(* IEC 61131-3 sources: JingjiangArm/moonboxpro_arm_8.4/Application/Application/任务列表/Main_Task/套色调整/套色新算法/PID_GET, 9 files *)

(* ---- AntiNotch_1.st ---- *)
(*@CES
Name=AntiNotch_1
Type=FunctionBlock
TypeGuid=6f9dac99-8de1-4efc-8465-68ac443b7d08
Guid=fc76d1c1-3b33-4f49-ab68-3746014dafce
HasDeclaration=True
HasImplementation=True
*)
{DECLARATION}
FUNCTION AntiNotch_1 : BOOL
(*功能：反陷波器(s^2+2*d*wn*s+wn^2)/(s^2+2*d*xi*wn*s+wn^2)的差分方程实现*)
(*输入：*)
(*输出：*)
VAR_INPUT
	i_rU:REAL;(*信号输入*)
	i_prYout: POINTER TO REAL;(*信号输出*)

(*(s^2+2*d*wn*s+wn^2)/(s^2+2*d*xi*wn*s+wn^2)*)
	i_rWn:REAL;(*陷波中心频率 rad/s*)
	i_rBw:REAL;(*陷波宽度 rad/s*)
	i_rDp:REAL;(*陷波深度 dB*)

	i_rTs:REAL;(*采样时间*)

	i_prUk:POINTER TO ARRAY [1..3] OF REAL;(*输入寄存器*)
	i_prYk:POINTER TO ARRAY [1..3] OF REAL;(*输出寄存器*)
END_VAR
VAR
	rFn:REAL:=0;
	rFBw:REAL:=0;
	rWn:REAL:=0;
	rDp:REAL:=0;

	rD:REAL:=0;
	rXi:REAL:=0;

	rK:REAL:=0;
	ra2:REAL:=0;
	ra1:REAL:=0;
	ra0:REAL:=0;

	rb2:REAL:=0;
	rb1:REAL:=0;
	rb0:REAL:=0;

	rTs:REAL:=0;(*采样时间*)
	rTemp:REAL:=0;

END_VAR
{IMPLEMENTATION}
(*参数初始化*)
rFn := i_rWn/2.0*gc_lrPi;
rWn := i_rWn;
rFBw := i_rBw/2.0*gc_lrPi;
rDp := i_rDp;

rTemp := -rDp/20.0;
rD := EXPT(10,rTemp);

rTemp := 1.0/(1.0 - 2.0*EXPT(rD,2));
rXi := rFBw/(2.0*rFn)*SQRT(rTemp);

rK := 1.0;

ra2:=1.0;
ra1:=2*rXi*rWn;
ra0:=rWn*rWn;

rb2:=1;
rb1:=2*rD*rXi*rWn;
rb0:=rWn*rWn;

rTs:=i_rTs;

(*更新寄存器注意顺序*)
i_prYk^[3]:=i_prYk^[2];
i_prYk^[2]:=i_prYk^[1];

i_prUk^[3]:=i_prUk^[2];
i_prUk^[2]:=i_prUk^[1];

(*差分计算*)
i_prUk^[1]:=rK*i_rU;
rTemp:=1/(rb0*rTs*rTs+2*rb1*rTs+4*rb2)*(-(2*rb0*rTs*rTs-8*rb2)*i_prYk^[2]-(rb0*rTs*rTs-2*rb1*rTs+4*rb2)*i_prYk^[3]
            +(ra0*rTs*rTs+2*ra1*rTs+4*ra2)*i_prUk^[1]+(2*ra0*rTs*rTs-8*ra2)*i_prUk^[2]+(ra0*rTs*rTs-2*ra1*rTs+4*ra2)*i_prUk^[3]);
i_prYk^[1]:=rTemp;
i_prYout^:=rTemp;

(* ---- Cal_Kp_Ki.st ---- *)
(*@CES
Name=Cal_Kp_Ki
Type=FunctionBlock
TypeGuid=6f9dac99-8de1-4efc-8465-68ac443b7d08
Guid=a93d564e-2599-4b4b-9c00-c963b5a75637
HasDeclaration=True
HasImplementation=True
*)
{DECLARATION}
FUNCTION Cal_Kp_Ki : BOOL
(*2024.9.6.123503*)
(*通过和控制器计算公式对比这里对Ki做的一些处理,反应到Ki计算上相当于积分的系数是定值,因为ts=周长/速度*系数
这里对输入的i_rV 按照30m/min定值输入,这样在计算积分的时候会出现积分根据速度逐渐减小的变化*)
(*2024.9.6.125139 将Ki的速度分开*)
(*2025.1.3.140421删除无用的*)
VAR_INPUT
(*
	i_byFilmType:BYTE;
	(*增加一些控制变量@2024.8.25.164242*)
	i_byTimingKiByArcErr:BYTE;(*=0 不使能|=1根据误差值Ki变化|值越大积分越小*)
	i_byAverageNum:BYTE;(*平均次数*)
	i_byColorId:BYTE;(*色序id*)
	i_iArcErr:INT;(*套色误差@mm*)
*)
(*模型变量*)
	i_rV:REAL;(*运行速度m/min*)
	i_rV_Ki:REAL;(*运行速度m/min*)
	i_rCL:REAL;(*版周长mm*)
	i_rL:REAL;(*机组料长m*)
(*控制变量*)
	i_rKadj_all:REAL;(*调整增益   40*)
	i_rKadj_i:REAL;(*积分增益  2.0*)
(*输出指针*)
	i_prKp:POINTER TO REAL;(*Kp*)
	i_prKi:POINTER TO REAL;(*Ki*)
END_VAR
VAR

	rA:REAL;(*模型参数*)(*
	iAverageNum:INT;
	iArcErr:INT;
*)
END_VAR
{IMPLEMENTATION}
IF i_rL<>0 AND i_rV<>0 AND i_rV_Ki<>0 AND i_rCL<>0 THEN
	(*计算模型参数*)
	rA := (i_rV/60.0)/i_rL;
	(*Kp*)
	i_prKp^ := i_rKadj_all/i_rCL*i_rV/rA;

	(*Ki*)
(*	i_prKi^ := i_rKadj_all/i_rCL*i_rV*i_rKadj_i;*)
	i_prKi^ := i_rKadj_all/i_rCL*i_rV_Ki*i_rKadj_i;
ELSE
	i_prKp^ := 16;
	i_prKi^ := 8;
END_IF

(* ---- Cal_Kp_Ki_V2.st ---- *)
(*@CES
Name=Cal_Kp_Ki_V2
Type=FunctionBlock
TypeGuid=6f9dac99-8de1-4efc-8465-68ac443b7d08
Guid=c47de549-0752-4bbe-8145-8113c580532b
HasDeclaration=True
HasImplementation=True
*)
{DECLARATION}
FUNCTION Cal_Kp_Ki_V2 : BOOL
(*2025.1.15.123422 增加了时延参数输入*)
VAR_INPUT
(*模型变量*)
	i_rV:REAL;(*运行速度m/min*)
	i_rLTao:REAL;(*印刷点到光电眼距离*)
	i_rL:REAL;(*机组料长m*)
	i_rDelay:REAL;(*时延@2025.1.15.123404+*)
(*控制变量*)
	i_rKadj_Mag:REAL;(*幅值裕度   15dB|越小越强*)
	i_rKadj_i:REAL;(*积分增益  1.0*)
(*输出指针*)
	i_prKp:POINTER TO REAL;(*Kp*)
	i_prKi:POINTER TO REAL;(*Ki*)
END_VAR
VAR
	rA:REAL;(*模型参数*)
	rTao:REAL;(*光电眼到印刷点的时延 s*)

	rWf:REAL;(*-180度对应的频率*)
	rMag_Wf:REAL;(*-180度对应的幅值*)

	rKadj:REAL; (*满足幅值裕度的增益*)
	rKTemp:REAL;(*增益计算临时变量*)

	iAverageNum:INT;
	iArcErr:INT;
END_VAR
{IMPLEMENTATION}
IF i_rL<>0 AND i_rV<>0 AND i_rLTao<>0 THEN
	(*计算模型参数*)
	rA := (i_rV/60.0)/i_rL;
(*	rTao := i_rLTao/(i_rV/60.0) +0.1 ;*)
	rTao := i_rLTao/(i_rV/60.0) + i_rDelay ;

	(*计算-180度对应的频率*)
	rWf := LREAL_TO_REAL(90.0 * gc_lrPi / 180.0 / rTao);
	(*计算-180度对应的幅值 和rKadj*)
	rMag_Wf := 20.0 * LOG(0.1 * rA / rWf); (*为负数*)
	rKTemp := (-1.0*i_rKadj_Mag - rMag_Wf) / 20.0  ;
	rKadj := LREAL_TO_REAL(EXPT(10, rKTemp));

	(*Kp*)
	i_prKp^ := rKadj;

	(*Ki*)
	i_prKi^ := rKadj * rA * i_rKadj_i;
ELSE
	i_prKp^ := 16;
	i_prKi^ := 8;
END_IF

(* ---- Cal_Kp_Ki_V3.st ---- *)
(*@CES
Name=Cal_Kp_Ki_V3
Type=FunctionBlock
TypeGuid=6f9dac99-8de1-4efc-8465-68ac443b7d08
Guid=deaeaf1e-1ab7-4a2c-8f0b-a36d361ddac8
HasDeclaration=True
HasImplementation=True
*)
{DECLARATION}
FUNCTION Cal_Kp_Ki_V3 : BOOL
(*2025.1.11.165519 增加了非法值处理@Liu.yt*)
(*将开环对象镇定为期望的幅值裕度和相位裕度*)
(*输入开环幅值裕度(10-20)，相位裕度(40-60)*)
(*由于需要调整积分满足相位裕度，因此实际的幅值裕度会略微小于设置值（在所给出的相位裕度范围内一般偏差在1dB以内，不超过2dB），相位裕度取得越小，幅值裕度偏差越大*)

VAR_INPUT
(*模型变量*)
	i_rV:REAL;(*运行速度m/min*)
	i_rLTao:REAL;(*印刷点到光电眼距离*)
	i_rL:REAL;(*机组料长m*)
(*控制变量*)
	i_rMargin_Mag:REAL;(*幅值裕度   15dB*)
	i_rMargin_Phi:REAL;(*相位裕度  50度*)
(*输出指针*)
	i_prKp:POINTER TO REAL;(*Kp*)
	i_prKi:POINTER TO REAL;(*Ki*)
END_VAR
VAR
	rA:REAL;(*模型参数*)
	rTao:REAL;(*光电眼到印刷点的时延 s*)

	rWf:REAL;(*-180度对应的频率*)
	rMag_Wf:REAL;(*-180度对应的幅值*)

	rKadj:REAL; (*满足幅值裕度的增益*)
	rKTemp:REAL;(*增益计算临时变量*)

	rKp_temp:REAL; (*临时Kp*)
	rKi_temp:REAL;(*临时Ki*)

	rax:REAL; (*模型临时参数，计算Wc使用*)
	rbx:REAL; (*模型临时参数，计算Wc使用*)

	rA_e:REAL;(*二次方程系数*)
	rB_e:REAL;(*二次方程系数*)
	rC_e:REAL;(*二次方程系数*)

	rX_temp:REAL;(*方程的解*)
	rWc:REAL;(*近似截止频率*)

	rPhi_temp:REAL;(*相位裕度临时量*)
	rDelta_Phi:REAL;(*相位裕度偏差*)
	rDelta_Phi_rad:REAL;(*相位裕度偏差 弧度表示*)

	rI:REAL;(*积分系数*)
END_VAR
{IMPLEMENTATION}
IF i_rL<>0 AND i_rV<>0 AND i_rLTao<>0 THEN
(*计算模型参数*)
	rA := (i_rV/60.0)/i_rL;
	rTao := i_rLTao/(i_rV/60.0) +0.1 ;
(*计算满足幅值裕度时的近似截止频率和增益*)
	(*计算-180度对应的频率*)
	rWf := LREAL_TO_REAL(90.0 * gc_lrPi / 180.0 / rTao);
	(*计算-180度对应的幅值 和rKadj*)
	rMag_Wf := 20.0 * LOG(0.1 * rA / rWf); (*为负数*)
	rKTemp := (-1.0*i_rMargin_Mag - rMag_Wf) / 20.0  ;
	rKadj := LREAL_TO_REAL(EXPT(10, rKTemp));

	(*Kp*)
	rKp_temp := rKadj;

	(*Ki*)
	rKi_temp := rKadj * rA;
	(*计算此时的截止频率Wc*)
	rax := rA;
	rbx := 0.1*rA;

	(*构建二次方程*)
	rA_e := 1;
	rB_e := rax * rax - rbx * rbx * rKp_temp * rKp_temp;
	rC_e := -1.0 * rbx * rbx * rKi_temp * rKi_temp;

	(*计算根*)
	rX_temp := (-1.0 * rB_e + SQRT(rB_e * rB_e - 4.0 * rA_e * rC_e)) / (2.0 * rA_e);
	rWc := SQRT(rX_temp);

	(*计算相位裕度偏差*)
	rPhi_temp := LREAL_TO_REAL(90.0 - rWc * rTao / gc_lrPi * 180.0);
	rDelta_Phi := rPhi_temp - i_rMargin_Phi - 5;(*5是额外的裕度，可调整*)

	rI := rA;
	IF rDelta_Phi > 0 THEN
		(*转成弧度表示*)
		rDelta_Phi_rad := LREAL_TO_REAL(rDelta_Phi / 180.0 * gc_lrPi);

		(*计算调整的积分系数rI *)
		rI := rWc * (1.0 + (rWc / rA) * TAN(rDelta_Phi_rad) ) /  ((rWc / rA) - TAN(rDelta_Phi_rad) );
	END_IF

	(*Kp*)
	i_prKp^ := rKadj;

	(*Ki*)
	i_prKi^ := rKadj * rI;
ELSE
	i_prKp^ := 16;
	i_prKi^ := 8;
END_IF

(* ---- Gc_Delta_PID_OutPut.st ---- *)
(*@CES
Name=Gc_Delta_PID_OutPut
Type=FunctionBlock
TypeGuid=6f9dac99-8de1-4efc-8465-68ac443b7d08
Guid=3bd2524c-3dcf-44dc-9cb0-138873b78811
HasDeclaration=True
HasImplementation=True
*)
{DECLARATION}
FUNCTION Gc_Delta_PID_OutPut : REAL
(*根据绝对值PID控制器输出和增量限幅计算实际的控制器输出增量*)
(*Input:绝对值PID控制器计算值 Cal_PID, 增量限幅值Limit_Delta, 当前控制量累计值*)
(*Output: 当前拍输出的控制量增量 Real_Delta_PID, 控制量累计值*)
VAR_INPUT
	i_rCal_PID:REAL;(*绝对值PID控制器计算值*)
	i_rLimit_Delta:REAL;(*增量限幅值 输入正值*)

	i_prReal_Delta_PID:POINTER TO REAL;(*当前拍输出的控制量增量*)
	i_prSigema_PID:POINTER TO REAL;(*控制量累计值*)
END_VAR

VAR
	rSigema_PID:REAL:=0.0;(*控制量累计值*)
	rGc_Delta:REAL:=0.0;(*当前绝对值PID输出与上一拍累计控制量的差*)
END_VAR
{IMPLEMENTATION}
(*内部变量赋值*)
rSigema_PID := i_prSigema_PID^;

(*计算当前绝对值PID输出与上一拍累计控制量的差*)
rGc_Delta := i_rCal_PID - rSigema_PID;

(*判断该差值的绝对值是否大于限幅值Limit_Delta*)
IF ABS(rGc_Delta) > i_rLimit_Delta THEN

	IF rGc_Delta >0 THEN
		i_prReal_Delta_PID^ := i_rLimit_Delta;
		i_prSigema_PID^ := rSigema_PID + i_rLimit_Delta;
	END_IF

	IF rGc_Delta <0 THEN
		i_prReal_Delta_PID^ := -i_rLimit_Delta;
		i_prSigema_PID^ := rSigema_PID - i_rLimit_Delta;
	END_IF

ELSE
	i_prReal_Delta_PID^ := rGc_Delta;
	i_prSigema_PID^ := rSigema_PID + rGc_Delta;
END_IF

(* ---- KS_GetPidParam.st ---- *)
(*@CES
Name=KS_GetPidParam
Type=FunctionBlock
TypeGuid=6f9dac99-8de1-4efc-8465-68ac443b7d08
Guid=5147df87-2533-411e-aab0-b9dfa23e86ce
HasDeclaration=True
HasImplementation=True
*)
{DECLARATION}
FUNCTION KS_GetPidParam : BOOL
(*2024.7.26.143250 重新调整*)
VAR_INPUT
	i_byFilmType: BYTE;
	i_byParamIndex: BYTE;
	(*以前的pid接口*)
	i_rKp_Hmi:REAL;
	i_rKi_Hmi:REAL;
	i_rKd_Hmi:REAL;
	i_rN_Hmi:REAL;

	(*模型输出的pid*)
	rKp_MolCal:REAL;
	rKi_MolCal:REAL;

	i_prKp: POINTER TO REAL;
	i_prKI: POINTER TO REAL;
	i_prKD: POINTER TO REAL;
	i_prN: POINTER TO REAL;
END_VAR
VAR
	rKp: REAL;
	rKI: REAL;
	rKD: REAL;
	rN: REAL;
END_VAR
{IMPLEMENTATION}
IF i_byParamIndex=1 THEN
	rKp:=16(*35*);
	rKI:=15(*2*);
	rKD:=0;
	rN:=0;
ELSIF i_byParamIndex=2 THEN
	rKp:=15.4634;
	rKI:=11.5601;
	rKD:=0;
	rN:=0;
ELSIF i_byParamIndex=3 THEN
	rKp:=17.3284;
	rKI:=6.0885;
	rKD:=0;
	rN:=0;
ELSIF i_byParamIndex=4 THEN
	rKp:=30;
	rKI:=0.3;
	rKD:=0;
	rN:=0;
ELSIF i_byParamIndex=9 THEN(*第9个参数作为模型pid*)
	rKp:=rKp_MolCal;
	rKI:=rKi_MolCal;
	rKD:=0;
	rN:=0;
ELSIF i_byParamIndex=10 THEN(*第10个参数作为手动输入的选择*)
	rKp:=i_rKp_Hmi;
	rKI:=i_rKi_Hmi;
	rKD:=i_rKd_Hmi;
	rN:=i_rN_Hmi;
ELSE
	rKp:=14.4215;
	rKI:=8.2591;
	rKD:=0;
	rN:=0;
END_IF

(*输出*)
IF i_prKp<>0 THEN
	i_prKp^:=rKp;
END_IF
IF i_prKI<>0 THEN
	i_prKI^:=rKI;
END_IF
IF i_prKd<>0 THEN
	i_prKd^:=rKD;
END_IF
IF i_prN<>0 THEN
	i_prN^:=rN;
END_IF

(* ---- Periodic.st ---- *)
(*@CES
Name=Periodic
Type=FunctionBlock
TypeGuid=6f9dac99-8de1-4efc-8465-68ac443b7d08
Guid=b9320914-a917-446b-b04f-68c6ab24df80
HasDeclaration=True
HasImplementation=True
*)
{DECLARATION}
FUNCTION Periodic : BOOL
(*自适应滤波器@频率要求特别准确*)
VAR_INPUT
(*输入输出*)
	i_rU:REAL;(*套色误差输入*)
	i_prYout: POINTER TO REAL;(*输出*)
(*
	i_prYout1: POINTER TO REAL;(*输出*)
	i_prYout2: POINTER TO REAL;(*输出*)
*)
(*系统参数*)
	i_rC:REAL;(*版周长mm*)
	i_rV:REAL;(*运行速度m/min*)
(*调整参数*)
	i_rG:REAL;(*趋近增益  不同频率可能符号改变*)
	i_rW:REAL;(*需要抑制的频率，应该尽可能精确*)

(*寄存器*)
	i_prTk:POINTER TO ARRAY [1..1] OF REAL;(*时间寄存器*)
	i_prTheta1k:POINTER TO ARRAY [1..1] OF REAL;(*Theta1寄存器*)
	i_prTheta2k:POINTER TO ARRAY [1..1] OF REAL;(*Theta2寄存器*)
END_VAR
VAR
(*模型参数*)
	rTs:REAL;

	rG:REAL;
	rW:REAL;

	rT:REAL;
	rTheta1:REAL;
	rTheta2:REAL;

	Dot_rTheta1:REAL;
	Dot_rTheta2:REAL;

	rTemp:REAL;
END_VAR
{IMPLEMENTATION}
(*参数初始化*)
	rTs := (i_rC/1000.0)/(i_rV/60.0);

	rG:=i_rG;
	rW:=i_rW;

	rT:=i_prTk^[1]*rTs;
	rTheta1:=i_prTheta1k^[1];
	rTheta2:=i_prTheta2k^[1];

(*计算*)
	Dot_rTheta1:=-1.0*rG*i_rU*COS(rW*rT);
	Dot_rTheta2:=-1.0*rG*i_rU*SIN(rW*rT);
rTemp:=rTheta1;
	rTheta1:=rTemp+Dot_rTheta1*rTs;
	rTheta2:=rTheta2+Dot_rTheta2*rTs;
(*输出*)
i_prYout^:=rTheta1*COS(rW*rT)+rTheta2*SIN(rW*rT);
(*
i_prYout1^:=rTheta1;
i_prYout2^:=rTheta2;
*)
(*寄存器更新*)
i_prTk^[1]:=i_prTk^[1]+1;
i_prTheta1k^[1]:=rTheta1;
i_prTheta2k^[1]:=rTheta2;

(* ---- Smith.st ---- *)
(*@CES
Name=Smith
Type=FunctionBlock
TypeGuid=6f9dac99-8de1-4efc-8465-68ac443b7d08
Guid=124e716f-cf6b-45b1-bef3-6a4f1ebc6f70
HasDeclaration=True
HasImplementation=True
*)
{DECLARATION}
FUNCTION Smith : BOOL
(*采取Smith的方法设计的控制器，只针对套色系统，采用滑动平均，长度3*)
(*平均次数不能随意修改@支持3幅平均*)
(*输入:*)
VAR_INPUT
(*输入输出*)
	i_rU:REAL;(*输入*)
	i_prYout: POINTER TO REAL;(*输出*)
(*系统参数*)
	i_rC:REAL;(*版周长mm*)
	i_rV:REAL;(*运行速度m/min*)
	i_rL:REAL;(*机组料长m*)
	i_iNDEL:INT;(*时延拍数N=LDel/C*)(*检测料长LDEL*)
(*寄存器  初始值0*)
(*0.1a/(s+a)*)
	i_prTF1Uk:POINTER TO ARRAY [1..2] OF REAL;(*输入寄存器*)
	i_prTF1Yk:POINTER TO ARRAY [1..2] OF REAL;(*输出寄存器*)
(*滑动滤波器(长度3) 1/3(z^2+z+1)/z^2*)
	i_prTF2Uk:POINTER TO ARRAY [1..3] OF REAL;(*输入寄存器*)
	i_prTF2Yk:POINTER TO ARRAY [1..3] OF REAL;(*输出寄存器*)
(*纯时延*)
	i_prDELUk:POINTER TO ARRAY [1..gc_iNDEL] OF REAL;(*输入寄存器*)

END_VAR

VAR
(*模型参数*)
	ra:REAL;
	rbc:REAL;

(*(a1s+a0)/(b1s+b0)*)
	rTF1IN:REAL;
	rTF1OUT:REAL;

	ra1_TF1:REAL;(*系统参数a1*)
	ra0_TF1:REAL;(*系统参数a0*)
	rb1_TF1:REAL;(*系统参数b1*)
	rb0_TF1:REAL;(*系统参数b0*)

(*(z^2+a1z+a0)/(z^2+b1z+b0)*)
	rTF2IN:REAL;
	rTF2OUT:REAL;

	ra2_TF2:REAL;(*系统参数a2*)
	ra1_TF2:REAL;(*系统参数a1*)
	ra0_TF2:REAL;(*系统参数a0*)
	rb2_TF2:REAL;(*系统参数b2*)
	rb1_TF2:REAL;(*系统参数b1*)
	rb0_TF2:REAL;(*系统参数b0*)

(*纯时延 *)
	iNDEL:INT;(*时延拍数*)
	rTF3IN:REAL;
	rTF3OUT:REAL;

	rTs:REAL:=0;(*采样时间*)
	rTemp:REAL:=0;

	iI:INT;(*循环拍数*)
END_VAR
{IMPLEMENTATION}
(*参数初始化*)
	ra := (i_rV/60.0)/i_rL;
	rbc := 0.1*ra;
	rTs := (i_rC/1000.0)/(i_rV/60.0);
(*TF1*)(*(a1s+a0)/(b1s+b0)*)
	rTF1IN := i_rU;

	ra1_TF1 := 0;(*a1*)
	ra0_TF1 := rbc;(*a0*)
	rb1_TF1 := 1.0;(*b1*)
	rb0_TF1 := ra;(*b0*)

	(*差分计算*)
	i_prTF1Uk^[1]:=rTF1IN;
	rTemp:=1.0/(rb0_TF1*rTs+2.0*rb1_TF1)*(-(rb0_TF1*rTs-2.0*rb1_TF1)*i_prTF1Yk^[2]+(ra0_TF1*rTs+2.0*ra1_TF1)*i_prTF1Uk^[1]+(ra0_TF1*rTs-2.0*ra1_TF1)*i_prTF1Uk^[2]);
	i_prTF1Yk^[1]:=rTemp;

	(*更新寄存器注意顺序*)
	i_prTF1Yk^[2]:=i_prTF1Yk^[1];
	i_prTF1Uk^[2]:=i_prTF1Uk^[1];

	rTF1OUT := i_prTF1Yk^[1];

(*TF2*)(*(a2z^2+a1z+a0)/(b2z^2+b1z+b0)*)
	rTF2IN := rTF1OUT;

	ra2_TF2:=1.0/3.0;(*a2*)
	ra1_TF2:=1.0/3.0;(*a1*)
	ra0_TF2:=1.0/3.0;(*a0*)
	rb2_TF2:=1.0;(*b2*)
	rb1_TF2:=0;(*b1*)
	rb0_TF2:=0;(*b0*)

	(*差分计算*)
	i_prTF2Uk^[1]:=rTF2IN;
	rTemp:=1.0/rb2_TF2*(-rb1_TF2*i_prTF2Yk^[2]-rb0_TF2*i_prTF2Yk^[3]+ra2_TF2*i_prTF2Uk^[1]+ra1_TF2*i_prTF2Uk^[2]+ra0_TF2*i_prTF2Uk^[3]);
	i_prTF2Yk^[1]:=rTemp;

	(*更新寄存器注意顺序*)
	i_prTF2Yk^[3]:=i_prTF2Yk^[2];
	i_prTF2Yk^[2]:=i_prTF2Yk^[1];

	i_prTF2Uk^[3]:=i_prTF2Uk^[2];
	i_prTF2Uk^[2]:=i_prTF2Uk^[1];

	rTF2OUT:=i_prTF2Yk^[1];

(*时延*)(*1-e^(ts)*)
	iNDEL := i_iNDEL;
(*差分计算*)
	rTF3IN:=rTF2OUT;
(*输出*)
	rTemp:=i_prDELUk^[iNDEL];
	i_prDELUk^[1]:=rTF3IN;
(*更新寄存器注意顺序*)
FOR iI:=0 TO iNDEL-2 BY 1 DO
	i_prDELUk^[iNDEL-iI]:=i_prDELUk^[iNDEL-iI-1];
END_FOR

rTF3OUT := rTF3IN-rTemp;
i_prYout^ := rTF3OUT;

(* ---- SmithPI.st ---- *)
(*@CES
Name=SmithPI
Type=FunctionBlock
TypeGuid=6f9dac99-8de1-4efc-8465-68ac443b7d08
Guid=cdff3448-9cdd-43dc-a40d-d24eec630f60
HasDeclaration=True
HasImplementation=True
*)
{DECLARATION}
FUNCTION SmithPI : BOOL
(*采取Smith的方法设计的控制器，只针对套色系统，采用滑动平均，长度3*)
(*输入:*)
VAR_INPUT
(*输入输出*)
	i_rU:REAL;(*输入*)
	i_prYout: POINTER TO REAL;(*输出*)
(*系统参数*)
	i_rC:REAL;(*版周长mm*)
	i_rV:REAL;(*运行速度m/min*)
	i_rL:REAL;(*机组料长m*)
	i_iNDEL:INT;(*时延拍数N=LDel/C*)(*检测料长LDEL*)
(*PI控制器*)
	i_rKp:REAL;(*版周长mm*)
	i_rKi:REAL;(*运行速度m/min*)
(*寄存器  初始值0*)
	i_prPIUk:POINTER TO ARRAY [1..2] OF REAL;(*输入寄存器*)
	i_prPIYk:POINTER TO ARRAY [1..2] OF REAL;(*输出寄存器*)
(*0.1a/(s+a)*)
	i_prTF1Uk:POINTER TO ARRAY [1..2] OF REAL;(*输入寄存器*)
	i_prTF1Yk:POINTER TO ARRAY [1..2] OF REAL;(*输出寄存器*)
(*滑动滤波器(长度3) 1/3(z^2+z+1)/z^2*)
	i_prTF2Uk:POINTER TO ARRAY [1..3] OF REAL;(*输入寄存器*)
	i_prTF2Yk:POINTER TO ARRAY [1..3] OF REAL;(*输出寄存器*)
(*纯时延*)
	i_prDELUk:POINTER TO ARRAY [1..gc_iNDEL] OF REAL;(*输入寄存器*)

END_VAR

VAR
(*模型参数*)
	ra:REAL;
	rbc:REAL;
(*PI*)
	rPIIN:REAL;
	rPIOUT:REAL;
	rKp:REAL;
	rKi:REAL;

(*(a1s+a0)/(b1s+b0)*)
	rTF1IN:REAL;
	rTF1OUT:REAL;

	ra1_TF1:REAL;(*系统参数a1*)
	ra0_TF1:REAL;(*系统参数a0*)
	rb1_TF1:REAL;(*系统参数b1*)
	rb0_TF1:REAL;(*系统参数b0*)

(*(z^2+a1z+a0)/(z^2+b1z+b0)*)
	rTF2IN:REAL;
	rTF2OUT:REAL;

	ra2_TF2:REAL;(*系统参数a2*)
	ra1_TF2:REAL;(*系统参数a1*)
	ra0_TF2:REAL;(*系统参数a0*)
	rb2_TF2:REAL;(*系统参数b2*)
	rb1_TF2:REAL;(*系统参数b1*)
	rb0_TF2:REAL;(*系统参数b0*)

(*纯时延 *)
	iNDEL:INT;(*时延拍数*)
	rTF3IN:REAL;
	rTF3OUT:REAL;

	rTs:REAL:=0;(*采样时间*)
	rTemp:REAL:=0;

	iI:INT;(*循环拍数*)
END_VAR
{IMPLEMENTATION}
(*参数初始化*)
	ra := (i_rV/60.0)/i_rL;
	rbc := 0.1*ra;
	rTs := (i_rC/1000.0)/(i_rV/60.0);
(*PI*)
	rKp:=i_rKp;
	rKi:=i_rKi;

	rTF2OUT:=i_prTF2Yk^[1];
	rPIIN:=i_rU-rTF2OUT;

	(*计算*)
	i_prPIUk^[1]:=rPIIN;
	i_prPIYk^[1]:=rKp*i_prPIUk^[1]+rTs*rKi*i_prPIYk^[2];
	(*更新寄存器注意顺序*)
	i_prPIYk^[2]:=i_prPIYk^[2]+i_prPIUk^[1];
	i_prPIUk^[2]:=i_prPIUk^[1];

	rPIOUT:=i_prPIYk^[1];
	i_prYout^:=rPIOUT;

(*TF1*)(*(a1s+a0)/(b1s+b0)*)
	rTF1IN := rPIOUT;

	ra1_TF1 := 0;(*a1*)
	ra0_TF1 := rbc;(*a0*)
	rb1_TF1 := 1.0;(*b1*)
	rb0_TF1 := ra;(*b0*)

	(*差分计算*)
	i_prTF1Uk^[1]:=rTF1IN;
	rTemp:=1.0/(rb0_TF1*rTs+2.0*rb1_TF1)*(-(rb0_TF1*rTs-2.0*rb1_TF1)*i_prTF1Yk^[2]+(ra0_TF1*rTs+2.0*ra1_TF1)*i_prTF1Uk^[1]+(ra0_TF1*rTs-2.0*ra1_TF1)*i_prTF1Uk^[2]);
	i_prTF1Yk^[1]:=rTemp;

	(*更新寄存器注意顺序*)
	i_prTF1Yk^[2]:=i_prTF1Yk^[1];
	i_prTF1Uk^[2]:=i_prTF1Uk^[1];

	rTF1OUT := i_prTF1Yk^[1];
(*时延*)(*1-e^(ts)*)
	iNDEL := i_iNDEL;
	(*差分计算*)
	rTF3IN:=rTF1OUT;
	(*输出*)
	rTemp:=i_prDELUk^[iNDEL];
	i_prDELUk^[1]:=rTF3IN;
	(*更新寄存器注意顺序*)
	FOR iI:=0 TO iNDEL-2 BY 1 DO
		i_prDELUk^[iNDEL-iI]:=i_prDELUk^[iNDEL-iI-1];
	END_FOR

	rTF3OUT := rTF3IN-rTemp;

(*TF2*)(*(z^2+a1z+a0)/(z^2+b1z+b0)*)
	rTF2IN := rTF3OUT;

	ra2_TF2:=1.0/3.0;(*a2*)
	ra1_TF2:=1.0/3.0;(*a1*)
	ra0_TF2:=1.0/3.0;(*a0*)
	rb2_TF2:=1.0;(*b2*)
	rb1_TF2:=0;(*b1*)
	rb0_TF2:=0;(*b0*)

	(*差分计算*)
	i_prTF2Uk^[1]:=rTF2IN;
	rTemp:=1.0/rb2_TF2*(-rb1_TF2*i_prTF2Yk^[2]-rb0_TF2*i_prTF2Yk^[3]+ra2_TF2*i_prTF2Uk^[1]+ra1_TF2*i_prTF2Uk^[2]+ra0_TF2*i_prTF2Uk^[3]);
	i_prTF2Yk^[1]:=rTemp;

	(*更新寄存器注意顺序*)
	i_prTF2Yk^[3]:=i_prTF2Yk^[2];
	i_prTF2Yk^[2]:=i_prTF2Yk^[1];

	i_prTF2Uk^[3]:=i_prTF2Uk^[2];
	i_prTF2Uk^[2]:=i_prTF2Uk^[1];
